{region 'Documentation'}
(*!
<summary>Check that IN is at most Maximum.</summary>
*)
{endregion}
FUNCTION_BLOCK AssertLessEqual_SInt EXTENDS AssertionBase
VAR_INPUT
    IN : SINT; //! Actual value checked or observed by this Assertion.
    Maximum : SINT; //! Inclusive upper bound of the comparison; for a range, must not be below Minimum.
END_VAR

SUPER^();

{region 'Documentation'}
(*!
<summary>Check that IN is at most Maximum.</summary>
*)
{endregion}
METHOD PROTECTED Assert
VAR
    Message : STRING(GVL_Constants.MessageLength);
    MaximumText : STRING(GVL_Constants.AssertionValueLength);
    ActualText : STRING(GVL_Constants.AssertionValueLength);
END_VAR
IF NOT EvaluationActive THEN
    RETURN;
END_IF;

IF Result = E_Result.Error THEN
    RETURN;
END_IF;

IF Result = E_Result.Failed THEN
    RETURN;
END_IF;

IF IN > Maximum THEN
    MaximumText := SINT_TO_STRING(Maximum);
    ActualText := SINT_TO_STRING(IN);
    Message := CONCAT('Assertion failed: value is above maximum. Maximum = ',
        MaximumText);
    Message := CONCAT(Message, ', Actual = ');
    Message := CONCAT(Message, ActualText);
    Message := CONCAT(Message, '.');
    Fail(Message := Message);
    RETURN;
END_IF;

Pass();
END_METHOD

END_FUNCTION_BLOCK

(* stored: Version 1.1.0.1
   POU AssertLessEqual_SInt: Id {9035e84a-289e-44e5-981d-ff92d74ee769}, SpecialFunc None
   Folder Internal: Id {00bdd251-de53-4254-a5be-cb423bba6313}
   Method Assert: Id {b685843c-827e-4d68-bfde-535a6bf2dfb0} *)
